Yaskawa INFORM job: -DEFRO-70_PRZYLACZE_60-DL40.JBI

/JOB
//NAME -DEFRO-70_PRZYLACZE_60-DL40
//POS
///NPOS 145,145,145,0,0,0
///TOOL 0
///POSTYPE PULSE
///PULSE
C00000=-281,-101163,-84214,3730,-80188,-1936
C00001=-283,-101162,-84213,3710,-80188,-1936
C00002=115939,-17843,-44700,-6904,-63515,59085
C00003=113314,-7643,-38017,-11019,-76954,88145
C00004=103027,16481,-40114,-5059,-61809,87383
C00005=105040,15326,-41057,-2867,-60895,82481
C00006=112116,-4038,-61231,4238,-38322,55452
C00007=119094,103,-60825,24445,-37916,40349
C00008=126451,21841,-45210,41120,-51782,12418
C00009=120810,45174,-18529,23033,-68771,15285
C00010=113661,48351,-10997,14394,-69817,-2320
C00011=99661,49426,-10503,-9214,-71488,-11368
C00012=100429,58976,-2984,-3175,-82283,-29084
C00013=89767,56609,-11491,-23507,-81851,-31378
C00014=90650,38781,-25820,-21905,-70921,-38459
C00015=94820,20520,-39102,-16125,-61441,-54226
C00016=98661,12402,-44932,-13704,-58284,-69648
C00017=98785,12241,-44972,-13685,-58324,-69693
C00018=99303,8604,-31154,-10952,-72489,-71699
C00019=89422,16015,-23794,-2157,-75183,91094
C00020=90147,29393,-27635,-2399,-65935,91035
C00021=95540,20095,-36882,3675,-57850,75382
C00022=103297,16374,-43607,17528,-50715,56089
C00023=113623,17176,-52780,50840,-45044,24405
C00024=112897,27423,-40548,43605,-50420,17252
C00025=110356,39314,-25385,32271,-59383,17432
C00026=104317,50857,-9144,20230,-66823,5878
C00027=93673,60339,2296,3658,-74232,-7297
C00028=87431,72964,12066,-3499,-86963,-24117
C00029=79200,70906,5432,-19177,-86971,-29152
C00030=76881,62048,-4360,-23768,-81676,-32231
C00031=75976,40412,-24595,-27810,-68313,-39866
C00032=79014,22952,-38581,-24432,-56090,-47051
C00033=83954,18821,-39545,-14696,-55602,-56766
C00034=84670,20170,-20597,-9101,-74704,-67115
C00035=72786,31521,-9549,-9445,-75352,93043
C00036=77700,39785,-17058,-2950,-63995,95472
C00037=81983,27857,-30062,1079,-52734,78101
C00038=87123,13822,-48367,12686,-33110,60100
C00039=91300,11273,-55373,33577,-24478,42822
C00040=99471,26612,-43555,50994,-41229,28947
C00041=98668,33324,-33405,41844,-45594,21473
C00042=97935,43024,-21733,40487,-51695,6645
C00043=90319,64223,7028,17469,-68688,4856
C00044=84028,80392,24912,7916,-81568,-6718
C00045=78609,83484,27340,-1219,-84898,-14295
C00046=77701,90823,33650,-789,-91896,-21073
C00047=70141,90423,29624,-15464,-93258,-27293
C00048=65818,68117,4765,-24481,-78068,-31304
C00049=68282,50646,-10447,-20317,-67064,-41748
C00050=69693,49887,-10181,-17194,-67455,-44679
C00051=70925,43946,-15385,-17448,-66914,-56829
C00052=75039,37514,-3449,-7701,-77257,-64173
C00053=74616,28156,-12897,-9694,-74827,92488
C00054=73831,40937,-16627,-11403,-64518,94085
C00055=79044,30924,-26494,-3857,-56066,85334
C00056=85009,15652,-44693,6448,-37732,65961
C00057=89198,10717,-53484,21981,-27493,50886
C00058=96896,19410,-49655,48443,-34236,32293
C00059=98470,33877,-32902,42106,-45617,19173
C00060=99425,42323,-24414,46724,-51265,3822
C00061=90043,63782,6675,17352,-68217,4924
C00062=76594,79956,24035,-8972,-81100,-4026
C00063=77844,90698,34010,-937,-91750,-20733
C00064=70407,90030,29268,-15583,-93200,-27364
C00065=66747,69510,6768,-22650,-79292,-32886
C00066=72490,51614,-6652,-10130,-69735,-47887
C00067=78982,35519,-21281,1001,-60006,-65808
C00068=74844,35432,-1015,-7610,-79822,-64270
C00069=74616,28156,-12897,-9694,-74827,92488
C00070=90411,-2677,-20047,-11125,-84138,86440
C00071=90413,-2674,-20051,-11105,-84138,86441
C00072=137757,-12075,-30464,2646,-72394,74401
C00073=139263,-65150,-85436,14259,-28990,73053
C00074=136879,-25803,-69250,35998,-11820,63023
C00075=139290,-23505,-65815,37849,-15870,40588
C00076=138255,-25667,-68923,45072,-10125,18948
C00077=137540,-11621,-49291,15825,-29065,282
C00078=134494,-8817,-45605,4069,-31945,-3289
C00079=134604,-8591,-45393,4272,-32069,-3452
C00080=134201,-22614,-63353,14441,-15462,-51172
C00081=133643,-21758,-61840,7774,-18256,-58833
C00082=132849,-22230,-62300,-146,-18489,-67744
C00083=134650,-26769,-71812,22381,-6082,-94556
C00084=132637,-74135,-100376,4983,-10333,-85647
C00085=119687,-78067,-87939,-2788,-20735,84624
C00086=119992,-27745,-68017,-3051,-15116,84333
C00087=119030,-28696,-69591,-21999,-13157,75803
C00088=119146,-27568,-67331,-20983,-14326,49763
C00089=119106,-25320,-64288,-16073,-16150,28459
C00090=116990,-27787,-67992,-36968,-13306,28443
C00091=114451,-20387,-59191,-34974,-24024,21051
C00092=114289,-23226,-63137,-42813,-20195,20855
C00093=115755,-27101,-67787,-45506,-13897,17108
C00094=116631,-28534,-69574,-43897,-10967,13052
C00095=119721,-30747,-72526,-5019,-4908,-12317
C00096=124673,-29524,-70968,54153,-12690,-50315
C00097=110381,-14519,-53439,-34713,-36084,-50985
C00098=115065,-20808,-58231,-19385,-28009,-64203
C00099=113126,-78683,-102705,-45607,-16425,-60367
C00100=120908,-77676,-80309,7462,-22023,84016
C00101=119355,-30092,-72700,-7480,-8883,86833
C00102=119330,-30666,-73900,-37441,-7256,75668
C00103=119392,-31005,-74194,-36731,-7285,75171
C00104=119107,-25533,-64139,-15884,-16345,28370
C00105=118189,-11113,-47154,-8478,-33276,7215
C00106=118285,-13415,-49709,-5227,-31034,-7778
C00107=112204,-14619,-53166,-28572,-30616,-12922
C00108=112459,-20642,-60567,-34495,-24493,-27463
C00109=113253,-23242,-63602,-34662,-21946,-37788
C00110=117822,-27208,-67860,-16762,-15410,-62087
C00111=114088,-29625,-74008,-62760,-13130,-51071
C00112=113074,-79856,-103225,-44998,-16651,-60643
C00113=120443,-70015,-86553,-1670,-18639,84017
C00114=119855,-29453,-70963,-4444,-11447,85360
C00115=119350,-27114,-66909,-10824,-16764,76179
C00116=120538,-28712,-69581,-9042,-12118,60389
C00117=121453,-23804,-62042,-1822,-20367,42740
C00118=119104,-25714,-64462,-15988,-16245,28420
C00119=118127,-25090,-63854,-17709,-16479,10287
C00120=118054,-20647,-58029,-8598,-22594,-6818
C00121=116391,-17852,-55102,-12391,-26715,-16410
C00122=113676,-17333,-55635,-24105,-28107,-26621
C00123=114148,-20487,-59353,-25400,-25301,-39443
C00124=114654,-26064,-67349,-36235,-17702,-47147
C00125=115014,-30497,-76060,-73901,-10838,-47744
C00126=112648,-89264,-107216,-40476,-18619,-62704
C00127=115490,-77010,-93554,-11224,-18305,89052
C00128=125433,-24819,-64014,25600,-22035,67229
C00129=124409,-21324,-58576,14136,-26697,62401
C00130=126029,-28427,-71429,47699,-12406,35561
C00131=126376,-14543,-51553,17453,-33391,37954
C00132=119104,-25707,-64456,-15987,-16243,28419
C00133=102227,-21803,-62565,-47260,-20333,28942
C00134=103256,-22698,-63333,-30550,-15064,8897
C00135=100032,-11798,-50575,-26640,-29993,-6479
C00136=97406,-10335,-50320,-35130,-33056,-18084
C00137=102127,-19671,-59474,-25169,-24074,-49644
C00138=96594,-22492,-70681,-79494,-21703,-41695
C00139=112538,-91654,-108181,-39431,-19159,-63177
C00140=113545,-73371,-70378,-16072,-42358,69017
C00141=89593,-90202,-78264,-12204,-55560,23671
C00142=60247,-88344,-77535,-12630,-64499,59028
C00143=11932,-100155,-87763,417,-74819,10359
C00144=-281,-101163,-84214,3730,-80188,-1936
BC00000=570125
BC00001=868704
BC00002=878894
BC00003=912823
BC00004=878035
BC00005=878036
BC00006=878037
BC00007=878037
BC00008=878037
BC00009=878038
BC00010=878038
BC00011=878037
BC00012=878037
BC00013=878037
BC00014=878037
BC00015=878037
BC00016=878037
BC00017=878037
BC00018=878037
BC00019=878035
BC00020=878036
BC00021=878037
BC00022=878037
BC00023=878038
BC00024=878038
BC00025=878038
BC00026=878038
BC00027=878037
BC00028=878037
BC00029=878037
BC00030=878037
BC00031=878037
BC00032=878037
BC00033=878037
BC00034=878037
BC00035=878037
BC00036=878035
BC00037=877203
BC00038=877947
BC00039=878201
BC00040=878342
BC00041=878784
BC00042=877962
BC00043=877604
BC00044=878141
BC00045=878500
BC00046=878840
BC00047=878535
BC00048=877975
BC00049=879348
BC00050=879174
BC00051=879174
BC00052=878037
BC00053=915550
BC00054=913919
BC00055=915607
BC00056=916395
BC00057=916456
BC00058=916387
BC00059=916442
BC00060=915550
BC00061=915870
BC00062=916359
BC00063=916876
BC00064=917058
BC00065=916344
BC00066=916666
BC00067=915811
BC00068=915811
BC00069=915550
BC00070=915550
BC00071=915550
BC00072=915550
BC00073=915550
BC00074=915550
BC00075=915550
BC00076=915550
BC00077=915550
BC00078=915550
BC00079=915550
BC00080=915550
BC00081=915550
BC00082=915550
BC00083=915550
BC00084=915550
BC00085=915550
BC00086=915551
BC00087=915550
BC00088=915550
BC00089=915550
BC00090=915550
BC00091=915550
BC00092=915550
BC00093=915550
BC00094=915550
BC00095=915550
BC00096=915550
BC00097=915550
BC00098=915550
BC00099=915550
BC00100=954211
BC00101=953187
BC00102=954162
BC00103=954160
BC00104=954071
BC00105=953684
BC00106=953455
BC00107=953244
BC00108=953665
BC00109=953702
BC00110=953799
BC00111=953749
BC00112=953683
BC00113=992214
BC00114=992214
BC00115=992103
BC00116=991968
BC00117=992423
BC00118=992186
BC00119=992082
BC00120=991590
BC00121=991168
BC00122=991569
BC00123=992150
BC00124=992735
BC00125=991845
BC00126=991844
BC00127=1026906
BC00128=1030289
BC00129=1030277
BC00130=1030261
BC00131=1030281
BC00132=1030485
BC00133=997557
BC00134=991657
BC00135=991168
BC00136=991569
BC00137=992735
BC00138=991845
BC00139=1030552
BC00140=1030552
BC00141=1015004
BC00142=995119
BC00143=847363
BC00144=570125
EC00000=1163,0
EC00001=1166,0
EC00002=-1742,0
EC00003=-1741,0
EC00004=-1745,0
EC00005=-1744,0
EC00006=-1742,0
EC00007=-1742,0
EC00008=-1741,0
EC00009=-1741,0
EC00010=-1741,0
EC00011=-1741,0
EC00012=-1741,0
EC00013=-1742,0
EC00014=-1742,0
EC00015=-1741,0
EC00016=-1741,0
EC00017=-1741,0
EC00018=-1741,0
EC00019=-1743,0
EC00020=-1742,0
EC00021=-1742,0
EC00022=-1742,0
EC00023=-1741,0
EC00024=-1741,0
EC00025=-1676,0
EC00026=-1724,0
EC00027=-1741,0
EC00028=-1741,0
EC00029=-1742,0
EC00030=-1742,0
EC00031=-1742,0
EC00032=-1742,0
EC00033=-1742,0
EC00034=-1741,0
EC00035=-1741,0
EC00036=-1743,0
EC00037=-1742,0
EC00038=-1743,0
EC00039=-1742,0
EC00040=-1741,0
EC00041=-1741,0
EC00042=-1741,0
EC00043=-1742,0
EC00044=-1741,0
EC00045=-1741,0
EC00046=-1741,0
EC00047=-1741,0
EC00048=-1741,0
EC00049=-1741,0
EC00050=-1741,0
EC00051=-1741,0
EC00052=-1741,0
EC00053=-1741,0
EC00054=-1742,0
EC00055=-1742,0
EC00056=-1743,0
EC00057=-1742,0
EC00058=-1741,0
EC00059=-1740,0
EC00060=-1741,0
EC00061=-1742,0
EC00062=-1742,0
EC00063=-1741,0
EC00064=-1741,0
EC00065=-1741,0
EC00066=-1742,0
EC00067=-1742,0
EC00068=-1741,0
EC00069=-1741,0
EC00070=-1741,0
EC00071=-84878,0
EC00072=-84879,0
EC00073=-84877,0
EC00074=-84877,0
EC00075=-84877,0
EC00076=-84877,0
EC00077=-84877,0
EC00078=-84877,0
EC00079=-84877,0
EC00080=-84877,0
EC00081=-84877,0
EC00082=-84877,0
EC00083=-84877,0
EC00084=-84877,0
EC00085=-84877,0
EC00086=-84878,0
EC00087=-84877,0
EC00088=-84877,0
EC00089=-84877,0
EC00090=-84877,0
EC00091=-84877,0
EC00092=-84877,0
EC00093=-84877,0
EC00094=-84877,0
EC00095=-84877,0
EC00096=-84877,0
EC00097=-84877,0
EC00098=-84877,0
EC00099=-84877,0
EC00100=-84877,0
EC00101=-84878,0
EC00102=-84877,0
EC00103=-84877,0
EC00104=-84877,0
EC00105=-84877,0
EC00106=-84877,0
EC00107=-84877,0
EC00108=-84877,0
EC00109=-84877,0
EC00110=-84877,0
EC00111=-84877,0
EC00112=-84877,0
EC00113=-84877,0
EC00114=-84877,0
EC00115=-84877,0
EC00116=-84877,0
EC00117=-84877,0
EC00118=-84877,0
EC00119=-84877,0
EC00120=-84877,0
EC00121=-84877,0
EC00122=-84877,0
EC00123=-84877,0
EC00124=-84877,0
EC00125=-84877,0
EC00126=-84877,0
EC00127=-84877,0
EC00128=-84877,0
EC00129=-84877,0
EC00130=-84877,0
EC00131=-84877,0
EC00132=-84877,0
EC00133=-84877,0
EC00134=-84877,0
EC00135=-84877,0
EC00136=-84877,0
EC00137=-84877,0
EC00138=-84877,0
EC00139=-84877,0
EC00140=-84877,0
EC00141=-1879,0
EC00142=-1342,0
EC00143=498,0
EC00144=1163,0
//INST
///DATE 2025/05/23 13:21
///COMM OZZ
///ATTR SC,RW
///GROUP1 RB1,BS1
///GROUP2 ST1
NOP
MOVJ C00000 BC00000 VJ=70.00 DEC=20  +MOVJ EC00000 VJ=70.00
MOVJ C00001 BC00001 VJ=40.00 DEC=20  +MOVJ EC00001 VJ=40.00
MOVJ C00002 BC00002 VJ=70.00 DEC=20  +MOVJ EC00002 VJ=70.00
MACRO1 MJ#(0) ARGF8
MOVJ C00003 BC00003 VJ=70.00 DEC=20  +MOVJ EC00003 VJ=0.78
MOVJ C00004 BC00004 VJ=80.00 DEC=20  +MOVJ EC00004 VJ=0.78
ARCON
MOVC C00005 BC00005 V=4.2 DEC=20  +MOVJ EC00005 VJ=0.78
MOVC C00006 BC00006 V=4.2 DEC=20  +MOVJ EC00006 VJ=30.00
MOVC C00007 BC00007 V=4.2 DEC=20  +MOVJ EC00007 VJ=30.00
MOVC C00008 BC00008 V=5.8 DEC=20  +MOVJ EC00008 VJ=30.00
MOVC C00009 BC00009 V=4.2 DEC=20  +MOVJ EC00009 VJ=30.00
MOVC C00010 BC00010 V=4.2 DEC=20  +MOVJ EC00010 VJ=30.00
MOVC C00011 BC00011 V=4.2 DEC=20  +MOVJ EC00011 VJ=30.00
MOVC C00012 BC00012 V=4.2 DEC=20  +MOVJ EC00012 VJ=30.00
MOVC C00013 BC00013 V=4.2 DEC=20  +MOVJ EC00013 VJ=30.00
MOVC C00014 BC00014 V=4.2 DEC=20  +MOVJ EC00014 VJ=30.00
MOVC C00015 BC00015 V=4.2 DEC=20  +MOVJ EC00015 VJ=30.00
MOVC C00016 BC00016 V=4.2 DEC=20  +MOVJ EC00016 VJ=30.00
MOVJ C00017 BC00017 VJ=25.00 DEC=20  +MOVJ EC00017 VJ=30.00
ARCOF
MOVJ C00018 BC00018 VJ=30.00 DEC=20  +MOVJ EC00018 VJ=30.00
MOVJ C00019 BC00019 VJ=30.00 DEC=20  +MOVJ EC00019 VJ=30.00
MOVJ C00020 BC00020 VJ=30.00 DEC=20  +MOVJ EC00020 VJ=30.00
ARCON
MOVC C00021 BC00021 V=4.2 DEC=20  +MOVJ EC00021 VJ=30.00
MOVC C00022 BC00022 V=4.2 DEC=20  +MOVJ EC00022 VJ=30.00
MOVC C00023 BC00023 V=4.2 DEC=20  +MOVJ EC00023 VJ=30.00
MOVC C00024 BC00024 V=4.2 DEC=20  +MOVJ EC00024 VJ=30.00
MOVC C00025 BC00025 V=4.2 DEC=20  +MOVJ EC00025 VJ=30.00
MOVC C00026 BC00026 V=4.2 DEC=20  +MOVJ EC00026 VJ=30.00
MOVC C00027 BC00027 V=4.2 DEC=20  +MOVJ EC00027 VJ=30.00
MOVC C00028 BC00028 V=4.2 DEC=20  +MOVJ EC00028 VJ=30.00
MOVC C00029 BC00029 V=4.2 DEC=20  +MOVJ EC00029 VJ=30.00
MOVC C00030 BC00030 V=4.2 DEC=20  +MOVJ EC00030 VJ=0.78
MOVC C00031 BC00031 V=5.8 DEC=20  +MOVJ EC00031 VJ=30.00
MOVC C00032 BC00032 V=4.2 DEC=20  +MOVJ EC00032 VJ=0.78
MOVC C00033 BC00033 V=4.2 DEC=20  +MOVJ EC00033 VJ=30.00
ARCOF
MOVJ C00034 BC00034 VJ=30.00 DEC=20  +MOVJ EC00034 VJ=30.00
MOVJ C00035 BC00035 VJ=30.00 DEC=20  +MOVJ EC00035 VJ=30.00
MOVJ C00036 BC00036 VJ=30.00 DEC=20  +MOVJ EC00036 VJ=30.00
ARCON
MOVC C00037 BC00037 V=4.2 DEC=20  +MOVJ EC00037 VJ=0.78
MOVC C00038 BC00038 V=4.2 DEC=20  +MOVJ EC00038 VJ=0.78
MOVC C00039 BC00039 V=4.2 DEC=20  +MOVJ EC00039 VJ=0.78
MOVC C00040 BC00040 V=4.2 DEC=20  +MOVJ EC00040 VJ=0.78
MOVC C00041 BC00041 V=4.2 DEC=20  +MOVJ EC00041 VJ=0.78
MOVC C00042 BC00042 V=4.2 DEC=20  +MOVJ EC00042 VJ=0.78
MOVC C00043 BC00043 V=4.2 DEC=20  +MOVJ EC00043 VJ=0.78
MOVL C00044 BC00044 V=4.2 DEC=20  +MOVJ EC00044 VJ=0.78
MOVC C00045 BC00045 V=4.2 DEC=20  +MOVJ EC00045 VJ=0.78
MOVC C00046 BC00046 V=4.2 DEC=20  +MOVJ EC00046 VJ=0.78
MOVC C00047 BC00047 V=4.2 DEC=20  +MOVJ EC00047 VJ=0.78
MOVC C00048 BC00048 V=4.2 DEC=20  +MOVJ EC00048 VJ=0.78
MOVC C00049 BC00049 V=4.2 DEC=20  +MOVJ EC00049 VJ=0.78
MOVC C00050 BC00050 V=4.2 DEC=20  +MOVJ EC00050 VJ=0.78
MOVC C00051 BC00051 V=4.2 DEC=20  +MOVJ EC00051 VJ=0.78
ARCOF
MOVJ C00052 BC00052 VJ=30.00 DEC=20  +MOVJ EC00052 VJ=30.00
MOVJ C00053 BC00053 VJ=30.00 DEC=20  +MOVJ EC00053 VJ=30.00
MOVJ C00054 BC00054 VJ=30.00 DEC=20  +MOVJ EC00054 VJ=30.00
ARCON
MOVC C00055 BC00055 V=4.2 DEC=20  +MOVJ EC00055 VJ=30.00
MOVC C00056 BC00056 V=4.2 DEC=20  +MOVJ EC00056 VJ=30.00
MOVC C00057 BC00057 V=4.2 DEC=20  +MOVJ EC00057 VJ=40.00
MOVC C00058 BC00058 V=4.2 DEC=20  +MOVJ EC00058 VJ=30.00
MOVC C00059 BC00059 V=4.2 DEC=20  +MOVJ EC00059 VJ=25.00
MOVC C00060 BC00060 V=4.2 DEC=20  +MOVJ EC00060 VJ=30.00
MOVC C00061 BC00061 V=4.2 DEC=20  +MOVJ EC00061 VJ=70.00
MOVC C00062 BC00062 V=4.2 DEC=20  +MOVJ EC00062 VJ=30.00
MOVC C00063 BC00063 V=4.2 DEC=20  +MOVJ EC00063 VJ=30.00
MOVC C00064 BC00064 V=4.2 DEC=20  +MOVJ EC00064 VJ=30.00
MOVC C00065 BC00065 V=4.2 DEC=20  +MOVJ EC00065 VJ=30.00
MOVC C00066 BC00066 V=4.2 DEC=20  +MOVJ EC00066 VJ=0.78
MOVC C00067 BC00067 V=4.2 DEC=20  +MOVJ EC00067 VJ=30.00
ARCOF
MOVJ C00068 BC00068 VJ=30.00 DEC=20  +MOVJ EC00068 VJ=30.00
MOVJ C00069 BC00069 VJ=30.00 DEC=20  +MOVJ EC00069 VJ=30.00
MOVJ C00070 BC00070 VJ=30.00 DEC=20  +MOVJ EC00070 VJ=30.00
MOVJ C00071 BC00071 VJ=30.00 DEC=20  +MOVJ EC00071 VJ=30.00
MOVJ C00072 BC00072 VJ=30.00 DEC=20  +MOVJ EC00072 VJ=30.00
MOVJ C00073 BC00073 VJ=70.00 DEC=20  +MOVJ EC00073 VJ=0.78
MOVJ C00074 BC00074 VJ=30.00 DEC=20  +MOVJ EC00074 VJ=0.78
MACRO1 MJ#(0) ARGF4
ARCON
MOVC C00075 BC00075 V=5.0 DEC=20  +MOVJ EC00075 VJ=0.78
MOVC C00076 BC00076 V=5.0 DEC=20  +MOVJ EC00076 VJ=0.78
MOVC C00077 BC00077 V=5.0 DEC=20  +MOVJ EC00077 VJ=0.78
MOVC C00078 BC00078 V=5.0 DEC=20  +MOVJ EC00078 VJ=0.78
MOVC C00079 BC00079 V=5.0 DEC=20  +MOVJ EC00079 VJ=0.78
MOVC C00080 BC00080 V=5.0 DEC=20  +MOVJ EC00080 VJ=0.78
MOVC C00081 BC00081 V=5.0 DEC=20  +MOVJ EC00081 VJ=0.78
MOVC C00082 BC00082 V=5.0 DEC=20  +MOVJ EC00082 VJ=0.78
MOVC C00083 BC00083 V=5.0 DEC=20  +MOVJ EC00083 VJ=0.78
ARCOF
MOVJ C00084 BC00084 VJ=40.00 DEC=20  +MOVJ EC00084 VJ=0.78
MOVJ C00085 BC00085 VJ=40.00 DEC=20  +MOVJ EC00085 VJ=0.78
MOVJ C00086 BC00086 VJ=40.00 DEC=20  +MOVJ EC00086 VJ=0.78
ARCON
MOVC C00087 BC00087 V=5.0 DEC=20  +MOVJ EC00087 VJ=0.78
MOVC C00088 BC00088 V=5.0 DEC=20  +MOVJ EC00088 VJ=40.00
MOVC C00089 BC00089 V=5.0 DEC=20  +MOVJ EC00089 VJ=0.78
MOVC C00090 BC00090 V=5.0 DEC=20  +MOVJ EC00090 VJ=0.78
MOVC C00091 BC00091 V=5.0 DEC=20  +MOVJ EC00091 VJ=0.78
MOVC C00092 BC00092 V=5.0 DEC=20  +MOVJ EC00092 VJ=0.78
MOVL C00093 BC00093 V=5.0 DEC=20  +MOVJ EC00093 VJ=80.00
MOVC C00094 BC00094 V=5.0 DEC=20  +MOVJ EC00094 VJ=0.78
MOVC C00095 BC00095 V=5.0 DEC=20  +MOVJ EC00095 VJ=0.78
MOVC C00096 BC00096 V=5.0 DEC=20  +MOVJ EC00096 VJ=0.78
MOVC C00097 BC00097 V=5.0 DEC=20  +MOVJ EC00097 VJ=70.00
MOVC C00098 BC00098 V=5.0 DEC=20  +MOVJ EC00098 VJ=0.78
ARCOF
MOVJ C00099 BC00099 VJ=40.00 DEC=20  +MOVJ EC00099 VJ=0.78
MOVJ C00100 BC00100 VJ=40.00 DEC=20  +MOVJ EC00100 VJ=0.78
MOVJ C00101 BC00101 VJ=40.00 DEC=20  +MOVJ EC00101 VJ=0.78
ARCON
MOVC C00102 BC00102 V=5.0 DEC=20  +MOVJ EC00102 VJ=0.78
MOVC C00103 BC00103 V=5.0 DEC=20  +MOVJ EC00103 VJ=0.78
MOVC C00104 BC00104 V=5.0 DEC=20  +MOVJ EC00104 VJ=0.78
MOVC C00105 BC00105 V=5.0 DEC=20  +MOVJ EC00105 VJ=0.78
MOVC C00106 BC00106 V=5.0 DEC=20  +MOVJ EC00106 VJ=0.78
MOVC C00107 BC00107 V=5.0 DEC=20  +MOVJ EC00107 VJ=0.78
MOVC C00108 BC00108 V=5.0 DEC=20  +MOVJ EC00108 VJ=0.78
MOVC C00109 BC00109 V=5.0 DEC=20  +MOVJ EC00109 VJ=0.78
MOVC C00110 BC00110 V=5.0 DEC=20  +MOVJ EC00110 VJ=0.78
MOVC C00111 BC00111 V=5.0 DEC=20  +MOVJ EC00111 VJ=0.78
ARCOF
MOVJ C00112 BC00112 VJ=40.00 DEC=20  +MOVJ EC00112 VJ=0.78
MOVJ C00113 BC00113 VJ=40.00 DEC=20  +MOVJ EC00113 VJ=0.78
MOVJ C00114 BC00114 VJ=40.00 DEC=20  +MOVJ EC00114 VJ=0.78
ARCON
MOVC C00115 BC00115 V=5.0 DEC=20  +MOVJ EC00115 VJ=0.78
MOVC C00116 BC00116 V=5.0 DEC=20  +MOVJ EC00116 VJ=0.78
MOVC C00117 BC00117 V=5.0 DEC=20  +MOVJ EC00117 VJ=0.78
MOVC C00118 BC00118 V=5.0 DEC=20  +MOVJ EC00118 VJ=0.78
MOVC C00119 BC00119 V=5.0 DEC=20  +MOVJ EC00119 VJ=0.78
MOVC C00120 BC00120 V=5.0 DEC=20  +MOVJ EC00120 VJ=0.78
MOVC C00121 BC00121 V=5.0 DEC=20  +MOVJ EC00121 VJ=0.78
MOVC C00122 BC00122 V=5.0 DEC=20  +MOVJ EC00122 VJ=0.78
MOVC C00123 BC00123 V=5.0 DEC=20  +MOVJ EC00123 VJ=0.78
MOVC C00124 BC00124 V=5.0 DEC=20  +MOVJ EC00124 VJ=0.78
MOVC C00125 BC00125 V=5.0 DEC=20  +MOVJ EC00125 VJ=0.78
ARCOF
MOVJ C00126 BC00126 VJ=40.00 DEC=20  +MOVJ EC00126 VJ=0.78
MOVJ C00127 BC00127 VJ=40.00 DEC=20  +MOVJ EC00127 VJ=0.78
MOVJ C00128 BC00128 VJ=40.00 DEC=20  +MOVJ EC00128 VJ=0.78
ARCON
MOVC C00129 BC00129 V=5.0 DEC=20  +MOVJ EC00129 VJ=0.78
MOVC C00130 BC00130 V=5.0 DEC=20  +MOVJ EC00130 VJ=0.78
MOVC C00131 BC00131 V=5.0 DEC=20  +MOVJ EC00131 VJ=0.78
MOVC C00132 BC00132 V=5.0 DEC=20  +MOVJ EC00132 VJ=0.78
MOVC C00133 BC00133 V=5.0 DEC=20  +MOVJ EC00133 VJ=70.00
MOVC C00134 BC00134 V=5.0 DEC=20  +MOVJ EC00134 VJ=30.00
MOVC C00135 BC00135 V=5.0 DEC=20  +MOVJ EC00135 VJ=70.00
MOVC C00136 BC00136 V=5.0 DEC=20  +MOVJ EC00136 VJ=70.00
MOVC C00137 BC00137 V=5.0 DEC=20  +MOVJ EC00137 VJ=70.00
MOVC C00138 BC00138 V=5.0 DEC=20  +MOVJ EC00138 VJ=70.00
ARCOF
MOVJ C00139 BC00139 VJ=40.00 DEC=20  +MOVJ EC00139 VJ=0.78
MOVJ C00140 BC00140 VJ=40.00 DEC=20  +MOVJ EC00140 VJ=0.78
MOVJ C00141 BC00141 VJ=40.00 DEC=20  +MOVJ EC00141 VJ=40.00
MOVJ C00142 BC00142 VJ=70.00 DEC=20  +MOVJ EC00142 VJ=0.78
MOVJ C00143 BC00143 VJ=70.00 DEC=20  +MOVJ EC00143 VJ=70.00
MOVJ C00144 BC00144 VJ=40.00 DEC=20  +MOVJ EC00144 VJ=0.78
END
